(* IEC 61131-3 sources: IRIS-Project/LASAL CONTROL SOFTWARE/LasalProject_2025_09_12/Class/_ModBusTCPSLAVE (part 2) *)

  pParameter := pData$^_ONE_ENTRY;                                                    // point to first entry of parameter list

  for i:=0 to (udEntryCount-1) do

    case pParameter^.usType of

      //=================================================================================
      MB_TYPE_SERVER: // parameter type ... server
      //=================================================================================
        if (pParameter^.ptr <> NIL) then                                                // is pointer valid ?
          pEntry^.ptr := pParameter^.ptr;                                               // add pointer to struct
        else
          retcode := MB_ERR_ADD_PARA;                                                   // set error code
          return;                                                                       // exit function because we do not handle with NILpointer
        end_if;

      //=================================================================================
      MB_TYPE_VARIABLE: // parameter type ... variable
      //=================================================================================
        if (pParameter^.ptr <> NIL) then                                                // is pointer valid ?
          pEntry^.ptr := pParameter^.ptr;                                               // add pointer to struct
        else                                                                            // invalid pointer
          retcode := MB_ERR_ADD_PARA;                                                   // set error code
          return;                                                                       // exit function because we do not handle with NILpointer
        end_if;

      //=================================================================================

    end_case;

    pEntry^.uiAddress := pParameter^.uiAddress;                                       // add MODBUS address to struct
    pEntry^.usReg     := pParameter^.usReg;                                           // add number of MODBUS register to struct
    pEntry^.usAccess  := pParameter^.usAccess;                                        // add parameter access rights to struct
    pEntry^.usType    := pParameter^.usType;                                          // add parameter type to struct
    pEntry^.dDataType := pParameter^.dDataType;                                       // add parameter data type to struct

    //----- type HOLDING registers  V.1.34 -----
    if (RegisterType = 0) then
      vAddrEntriesHolding.udNo += 1;                                                  // increase the number of entries
      pEntry^.udEntryNo := vAddrEntriesHolding.udNo;                                  // set the actual entry number
    end_if;
    //----- type INPUT registers  V.1.34 -----
    if (RegisterType = 1) then
      vAddrEntriesInput.udNo += 1;                                                    // increase the number of entries
      pEntry^.udEntryNo := vAddrEntriesInput.udNo;                                    // set the actual entry number
    end_if;

    pParameter += sizeof(_ONE_ENTRY);                                                 // point to next parameter
    pEntry     += sizeof(_ONE_ENTRY);                                                 // point to next free entry

  end_for;

  //----- type HOLDING registers  V.1.34 -----
  if (RegisterType = 0) then
    if (vAddrEntriesHolding.udNo < to_UDINT(cBufSize)) then                           // buffer isn't full
      pEntry += sizeof(_ONE_ENTRY);                                                   // set pointer to the next free space in allocated memory
      INIT_ENTRY(ptr:=pEntry);                                                        // clear the next space in allocated memory
    end_if;
  end_if;
  //----- type INPUT registers  V.1.34 -----
  if (RegisterType = 1) then
    if (vAddrEntriesInput.udNo < to_UDINT(cBufSizeInputReg)) then                     // buffer isn't full
      pEntry += sizeof(_ONE_ENTRY);                                                   // set pointer to the next free space in allocated memory
      INIT_ENTRY(ptr:=pEntry);                                                        // clear the next space in allocated memory
    end_if;
  end_if;

  SortEntries(RegisterType);

END_FUNCTION

FUNCTION VIRTUAL _ModBusTCPSLAVE::ExceptionLogging
VAR_INPUT
  pRequest 	      : ^_REQUEST;
  ExceptionCode 	: USINT;
END_VAR
VAR
	szLogEntry      : ARRAY [0..255] OF CHAR;
  dValue          : DINT;
  szValue         : ARRAY [0..15] OF CHAR;
  szHelp          : ARRAY [0..15] OF CHAR;
  udStrLen        : UDINT;
  i               : USINT;
END_VAR

  // -----------------------------------------------------------------
  // - ADD FUNCTION CODE TO LOG ENTRY
  // -----------------------------------------------------------------
  coSigCLib.StrCpy(#szLogEntry[0], "Modbus Slave Exception Response, Function=");
  dValue := to_DINT(pRequest^.usFunction);
  coSigCLib.IToA(dValue, #szValue[0], 10);
  coSigCLib.StrCat(#szLogEntry[0], #szValue[0]);
  // -----------------------------------------------------------------
  // - ADD EXCEPTION CODE TO LOG ENTRY
  // -----------------------------------------------------------------
  coSigCLib.StrCat(#szLogEntry[0], ", Exception Code=");
  dValue := to_DINT(ExceptionCode);
  coSigCLib.IToA(dValue, #szValue[0], 10);
  coSigCLib.StrCat(#szLogEntry[0], #szValue[0]);
  // -----------------------------------------------------------------
  // - ADD OBJECT ADDRESS TO LOG ENTRY
  // -----------------------------------------------------------------
  coSigCLib.StrCat(#szLogEntry[0], ", this=");
  coSigCLib.IToA(this$DINT, #szValue[0], 0x10);
  udStrLen := coSigCLib.StrLen(#szValue[0]);

  i := 2;
  szHelp[0] := '0';
  szHelp[1] := 'x';
  szHelp[2] := 0x00;

  while udStrLen < 0x08 do
    szHelp[i]   := '0';
    szHelp[i+1] := 0x00;
    udStrLen    += 1;
    i           += 1;
  end_while;

  coSigCLib.StrCat(#szHelp[0], #szValue[0]);
  coSigCLib.StrCat(#szLogEntry[0], #szHelp[0]);

  coSysMsg.ULPrintfln0(#szLogEntry[0]);

  ExceptionLoggingDetail(pRequest);

END_FUNCTION

FUNCTION VIRTUAL _ModBusTCPSLAVE::ExceptionLoggingDetail
VAR_INPUT
  pRequest 	: ^_REQUEST;
END_VAR
VAR
	szLogEntry    : ARRAY [0..255] OF CHAR;
  szValue       : ARRAY [0..15] OF CHAR;
  uiValue       : UINT;
END_VAR

  case pRequest^.usFunction of

    (*=======================================================================*)
    MB_FUNC_RD_MULTIPLE_REG:
    (*=======================================================================*)
      coSigCLib.StrCpy(#szLogEntry[0], "---Detailed Information: StartAddress=");
      if (cTurnBytes = 0) then
        uiValue := pRequest^.aData[0]$UINT;
      else
        uiValue := Turn_2_Bytes(pRequest^.aData[0]$UINT);
      end_if;
      coSigCLib.IToA(to_DINT(uiValue), #szValue[0], 10);
      coSigCLib.StrCat(#szLogEntry[0], #szValue[0]);
      coSigCLib.StrCat(#szLogEntry[0], ", RegisterCnt=");
      if (cTurnBytes = 0) then
        uiValue := pRequest^.aData[2]$UINT;
      else
        uiValue := Turn_2_Bytes(pRequest^.aData[2]$UINT);
      end_if;
      coSigCLib.IToA(to_DINT(uiValue), #szValue[0], 10);
      coSigCLib.StrCat(#szLogEntry[0], #szValue[0]);
      coSigCLib.StrCat(#szLogEntry[0], ", StartAddrOffset=");
      coSigCLib.IToA(StartAddrOffset, #szValue[0], 10);
      coSigCLib.StrCat(#szLogEntry[0], #szValue[0]);
      coSigCLib.StrCat(#szLogEntry[0], ", UseOffset=");
      coSigCLib.IToA(UseOffset, #szValue[0], 10);
      coSigCLib.StrCat(#szLogEntry[0], #szValue[0]);

      coSysMsg.ULPrintfln0(#szLogEntry[0]);

    (*=======================================================================*)
    MB_FUNC_RD_MULTIPLE_INPUT_REG:
    (*=======================================================================*)
      coSigCLib.StrCpy(#szLogEntry[0], "---Detailed Information: StartAddress=");
      if (cTurnBytes = 0) then
        uiValue := pRequest^.aData[0]$UINT;
      else
        uiValue := Turn_2_Bytes(pRequest^.aData[0]$UINT);
      end_if;
      coSigCLib.IToA(to_DINT(uiValue), #szValue[0], 10);
      coSigCLib.StrCat(#szLogEntry[0], #szValue[0]);
      coSigCLib.StrCat(#szLogEntry[0], ", RegisterCnt=");
      if (cTurnBytes = 0) then
        uiValue := pRequest^.aData[2]$UINT;
      else
        uiValue := Turn_2_Bytes(pRequest^.aData[2]$UINT);
      end_if;
      coSigCLib.IToA(to_DINT(uiValue), #szValue[0], 10);
      coSigCLib.StrCat(#szLogEntry[0], #szValue[0]);
      coSigCLib.StrCat(#szLogEntry[0], ", StartAddrOffsInputReg=");
      coSigCLib.IToA(StartAddrOffsInputReg, #szValue[0], 10);
      coSigCLib.StrCat(#szLogEntry[0], #szValue[0]);
      coSigCLib.StrCat(#szLogEntry[0], ", UseOffsInputReg=");
      coSigCLib.IToA(UseOffsInputReg, #szValue[0], 10);
      coSigCLib.StrCat(#szLogEntry[0], #szValue[0]);

      coSysMsg.ULPrintfln0(#szLogEntry[0]);

    (*=======================================================================*)
    MB_FUNC_WR_MULTIPLE_REG:
    (*=======================================================================*)
      coSigCLib.StrCpy(#szLogEntry[0], "---Detailed Information: StartAddress=");
      if (cTurnBytes = 0) then
        uiValue := pRequest^.aData[0]$UINT;
      else
        uiValue := Turn_2_Bytes(pRequest^.aData[0]$UINT);
      end_if;
      coSigCLib.IToA(to_DINT(uiValue), #szValue[0], 10);
      coSigCLib.StrCat(#szLogEntry[0], #szValue[0]);
      coSigCLib.StrCat(#szLogEntry[0], ", RegisterCnt=");
      if (cTurnBytes = 0) then
        uiValue := pRequest^.aData[2]$UINT;
      else
        uiValue := Turn_2_Bytes(pRequest^.aData[2]$UINT);
      end_if;
      coSigCLib.IToA(to_DINT(uiValue), #szValue[0], 10);
      coSigCLib.StrCat(#szLogEntry[0], #szValue[0]);
      coSigCLib.StrCat(#szLogEntry[0], ", StartAddrOffset=");
      coSigCLib.IToA(StartAddrOffset, #szValue[0], 10);
      coSigCLib.StrCat(#szLogEntry[0], #szValue[0]);
      coSigCLib.StrCat(#szLogEntry[0], ", UseOffset=");
      coSigCLib.IToA(UseOffset, #szValue[0], 10);
      coSigCLib.StrCat(#szLogEntry[0], #szValue[0]);

      coSysMsg.ULPrintfln0(#szLogEntry[0]);

  end_case;

END_FUNCTION
